(*
SPDX-FileCopyrightText: © 2026 Oleksandr Tiutyk <trofimich@gmail.com>
SPDX-License-Identifier: MIT
License: https://opensource.org/license/mit
*)

(*!
<summary>Provides finite bounds for UnsignedInt16 values.</summary>
<description>
MIN_VALUE and MAX_VALUE describe the represented integer range; constants perform no conversion or runtime
validation. Additional named bounds, where declared, describe narrower representations.
</description>
*)

{attribute 'no_explicit_call' := 'do not call this function block directly'}
PROGRAM UnsignedInt16
VAR CONSTANT
	ZERO : UINT := 0;
	MIN_VALUE : UINT := 0;
	MAX_VALUE : UINT := UINT#16#FFFF;
END_VAR
VAR
	{attribute 'hide'} 
	_ClassName : STRING := __POUNAME();
END_VAR

{attribute 'monitoring' := 'call'}
PROPERTY ClassName : REFERENCE TO STRING
GET
ClassName REF= _ClassName;
END_GET
END_PROPERTY

(*!
<summary>Provides the library namespace used in diagnostics.</summary>
<description>
Borrowed read-only reference to the compiler-initialized library namespace; no ownership transfer.
</description>
*)
{attribute 'monitoring' := 'call'}
PROPERTY NamespaceName : REFERENCE TO STRING
GET
NamespaceName REF= CurrentNamespace.Name;
END_GET
END_PROPERTY

END_PROGRAM

(* stored: Version 1.1.0.1
   POU UnsignedInt16: Id {359c1cce-ae3b-4104-951e-6498f593d0f2}, SpecialFunc None
   Property ClassName: Id {e28f3e6b-f8ef-4f8f-aaca-b868322c98eb}
   Get Get: Id {91af5dcb-ef23-4bee-8853-6d037edab072}
   Property NamespaceName: Id {de673b86-8af7-471b-8059-506452281cca}
   Get Get: Id {c5c97b87-3837-4e30-b5d4-b8fd59f60799} *)
